Fanuc KAREL source: kb00020.KL

-- PROVISIONAL review KL for V770-1; original PC SHA256 6276504d1581c7358a62abe6b283d7276da7ccde4257c0feec1f9eeb8ffa40a2
-- Incomplete behavior may be omitted. Consult companion uncertainty JSON. Do not deploy.
PROGRAM KB00020
%NOLOCKGROUP
VAR
  P1 : INTEGER
  RESULT : STRING[80]
BEGIN
  -- UNRESOLVED_PC offsets 5-12; opcodes 9D,23
  -- UNRESOLVED_PC offsets 17-32; opcodes 27,22,76,75
  -- UNRESOLVED_PC offsets 37-41; opcodes 7F
END KB00020
